SUBAPPLICATION Schneidwerk (* Subapplication Type *)
  (* Standard: 61499-2 *)
  (* Version 1.0, 2023-01-29, Franz *)
  IMPORT DefaultPool::SoftKey_Schneidwerk;
  IMPORT isobus::UT::io::Softkey::SoftKeyActivationCode::SK_RELEASED;
  IMPORT DefaultPool::AuxInput_Schneidwerk;
  IMPORT isobus::UT::io::Auxiliary::IN::AuxiliaryState::AuxDisabled;
  IMPORT DataPanel::io::MI::DQ::DataPanel_MI_DO::DigitalOutput_1A;
  IMPORT DataPanel::io::MI::DQ::DataPanel_MI_DO::DigitalOutput_1B;
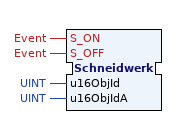
  EVENT_INPUT
    S_ON;
    S_OFF;
  END_EVENT
  VAR_INPUT
    u16ObjId : UINT;
    u16ObjIdA : UINT;
  END_VAR
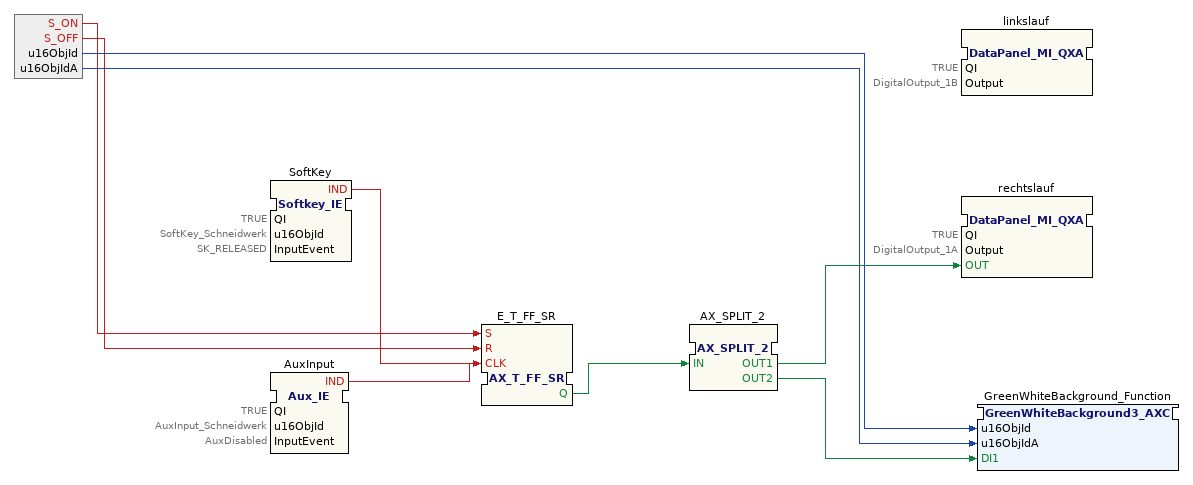
  (* TODO: Schneidwerk linkslauf bei jedem 2. Start. *)
  FBS
    rechtslauf : DataPanel::io::MI::DQ::DataPanel_MI_QXA(QI := TRUE, Output := DigitalOutput_1A);
    E_T_FF_SR : adapter::events::unidirectional::AX_T_FF_SR;
    AX_SPLIT_2 : adapter::events::unidirectional::AX_SPLIT_2;
    linkslauf : DataPanel::io::MI::DQ::DataPanel_MI_QXA(QI := TRUE, Output := DigitalOutput_1B);
    SoftKey : isobus::UT::io::Softkey::Softkey_IE(QI := TRUE, u16ObjId := SoftKey_Schneidwerk, InputEvent := SK_RELEASED);
    AuxInput : isobus::UT::io::Auxiliary::IN::Aux_IE(QI := TRUE, u16ObjId := AuxInput_Schneidwerk, InputEvent := AuxDisabled);
  END_FBS
  SUBAPPS
    GreenWhiteBackground_Function : MyLib::sys::GreenWhiteBackground3_AXC;
  END_SUBAPPS
  EVENT_CONNECTIONS
    S_ON TO E_T_FF_SR.S;
    S_OFF TO E_T_FF_SR.R;
    SoftKey.IND TO E_T_FF_SR.CLK;
    AuxInput.IND TO E_T_FF_SR.CLK;
  END_CONNECTIONS
  DATA_CONNECTIONS
    u16ObjId TO GreenWhiteBackground_Function.u16ObjId;
    u16ObjIdA TO GreenWhiteBackground_Function.u16ObjIdA;
  END_CONNECTIONS
  ADAPTER_CONNECTIONS
    E_T_FF_SR.Q TO AX_SPLIT_2.IN;
    AX_SPLIT_2.OUT1 TO rechtslauf.OUT;
    AX_SPLIT_2.OUT2 TO GreenWhiteBackground_Function.DI1;
  END_CONNECTIONS
END_SUBAPPLICATION
